// Communication API/Ethernet/API/bds_ethIPv4_setLocalIpAdr
///This function sets the IPv4 Address and Subnet Mask of the ECU.
///
///=======
/// Remarks:
///=======
///This function must be called from initialization task. 
///IP address shall be Unicast only. Multicast (from 0xE0000000 to 0xEFFFFFFF) or broadcast (0xFFFFFFFF) or 0 are not allowed.
///The Subnet mask(CIDR) can have any value from 1 to 31.
///If this API is called properly from OsIniProc(), then it will overwrite the IP address configured in easyConfig.
///The header file bds_ethIPv4_SetIPAdr.h shall be included for enabling usage of defines.
///----------
/// FFI:
///----------
///This API can be used in trusted partitions only. See Freedom from Interference (FFI) concept for more details.
///
///==================================================================		  	===================================================================================================
///Return value    								  							    Description
///==================================================================		  	===================================================================================================
///bds_ethIPv4_Adr_Mask_ok_E                                                    API call is successful
///bds_ethIPv4_Adr_Nok_E                                                        API call is invalid because of invalid IPv4 address, Unicast address expected.
///bds_ethIPv4_Mask_Nok_E 	                                                    API call is invalid because of invalid subnet mask, subnet mask should be 16.
///bds_ethIPv4_Api_NotAvailable_E                                               Not Available (e.g. busy, called too early in init, not called from OsIniProc etc.)
///
///==================================================================		   	===================================================================================================
///=======
///Code Example:
///=======
/// PROGRAM ETHERNET
/// VAR
///   bds_ethIPv4_Set_Adr_Mask_s1 : bds_ethIPv4_LocalIpAdr_ts;
///   flag_u8 : USINT := 0;
/// END_VAR
///
/// (* Set IP Address: 192.168.0.3 (0xC0A80003) *)
/// bds_ethIPv4_Set_Adr_Mask_s1.Ipv4Adr_u32 := 16#C0A80003; 
///
/// (* Set Subnet Mask: /16 (255.255.0.0) *)
/// bds_ethIPv4_Set_Adr_Mask_s1.Ipv4SubnetMask_u8 := 16;
///
/// (* Apply IP configuration *)
/// 
/// IF(flag_u8 = 0) THEN
/// bds_ethIPv4_setLocalIpAdr(bds_ethIPv4_Set_Adr_Mask_s1);
///
/// flag_u8 :=1;
/// END_IF
/// END_PROGRAM
///============================================================================
{attribute 'external_name' := 'cmp_rts_bds_ethIPv4_setLocalIpAdr'}
FUNCTION bds_ethIPv4_setLocalIpAdr : bds_ethIPv4_setLocalIpAdr_ts
VAR_INPUT
	//Data Structure for IPv4 Address and Subnet Mask
	bds_ethIPv4_setLocalIpAdr_s : bds_ethIPv4_LocalIpAdr_ts;
END_VAR

END_FUNCTION

// Communication API/Ethernet/API/bds_ethIPv4_getLocalIpAdr
///This function reads the IPv4 Address and Subnet Mask of the ECU.
///
///=======
/// Remarks:
///=======
///The header file bds_ethIPv4_SetIPAdr.h shall be included for enabling usage of defines.
///----------
/// FFI:
///----------
///This API can be used in trusted partitions only. See Freedom from Interference (FFI) concept for more details.
///
///==================================================================		  	===================================================================================================
///Return value    								  							    Description
///==================================================================		  	===================================================================================================
///bds_ethIPv4_Adr_Mask_ok_E                                                    API call is successful
///bds_ethIPv4_Api_NotAvailable_E                                               Not Available (e.g. busy, called too early in init, not called from OsIniProc etc.)
///bds_ethIPv4_NullPtr_E                                                        Invalid parameter passed
///==================================================================		   	===================================================================================================
///=======
///Code Example:
///=======
///PROGRAM ETHERNET
/// VAR
///    bds_ethIPv4_Get_Adr_Mask_s2 : bds_ethIPv4_LocalIpAdr_ts;
/// END_VAR
/// 
/// bds_ethIPv4_Get_Adr_Mask_s2.Ipv4Adr_u32 := 0;
/// bds_ethIPv4_Get_Adr_Mask_s2.Ipv4SubnetMask_u8 := 0;
///
/// bds_ethIPv4_getLocalIpAdr(ADR(bds_ethIPv4_Get_Adr_Mask_s2));
///
///END_PROGRAM
///============================================================================
{attribute 'external_name' := 'cmp_rts_bds_ethIPv4_getLocalIpAdr'}
FUNCTION bds_ethIPv4_getLocalIpAdr : bds_ethIPv4_getLocalIpAdr_ts
VAR_INPUT
	//Data Structure for IPv4 Address and Subnet Mask
	bds_ethIPv4_getLocalIpAdr_s : POINTER TO bds_ethIPv4_LocalIpAdr_ts;
END_VAR

END_FUNCTION

// Communication API/Ethernet/API/bds_ethIPv4_setDoipAdr
///This function configures the RC4x's and Tester's logical addresses for Diagnostic over IP (DoIP) communication. 
///
///=======
/// Remarks:
///=======
///This function shall be called from initialization task.
///The logical address of the RC4x (ecuLogAdr_u16) must fall within one of two valid ranges, as defined by ISO 13400-2:
/// Standard ECU addresses - 0x0001 to 0x0DFF
/// Extended ECU addresses - 0x1000 to 0x7FFF.
/// An address outside these ranges will result in bds_ethIPv4_retLogAdrNok_E.
///The Tester logical address (testerLogAdr_u16) must be within the range 0x0E00 to 0x0FFF. An address outside this range will result in bds_ethIPv4_retTesterAdrNok_E.
///If this API is not called, or called incorrectly (validation fails , bds_ethIPv4_retTesterAdrNok_E), the RC4x shall use the addresses from easyConfig.
///This function call overrides the statically configured values provided by easyConfig.
///----------
/// FFI:
///----------
///This API can be used in trusted partitions only. See Freedom from Interference (FFI) concept for more details.
///
///==================================================================		  	===================================================================================================
///Return value    								  							    Description
///==================================================================		  	===================================================================================================
///ecuLogAdr_u16                                                                API call is successful
///testerLogAdr_u16                                                             Tester logical address (valid range: 0x0E00-0x0FFF)
///
///==================================================================		   	===================================================================================================
///=======
///Code Example:
///=======
///PROGRAM ETHERNET
/// VAR
///    doipStatus : bds_ethIPv4_retDoipAdr_te;
///    flag_u8 : USINT := 0;
/// END_VAR

(* Configure ECU Logical Target Address and Tester Address Range
 *
 * ECU Logical Target Address = 0x0200
 * Tester Address Range Min   = 0x0E00
 *
 * NOTE: The Tester Address Range Max is internally defined in the stack.
 *)
/// IF(flag_u8 = 0) THEN
/// doipStatus := bds_ethIPv4_setDoipAdr(16#0200, 16#0E00);
/// 
/// flag_u8 := 1;
/// 
/// END_IF
///
(* Check return status *)
/// IF doipStatus = bds_ethIPv4_retAdrOk_E THEN
   (* DoIP address successfully configured*)
    
/// ELSE
    (* Error handling: DoIP address configuration failed*)
    
/// END_IF;

/// END_PROGRAM
///============================================================================
{attribute 'external_name' := 'cmp_rts_bds_ethIPv4_setDoipAdr'}
FUNCTION bds_ethIPv4_setDoipAdr : bds_ethIPv4_retDoipAdr_te
VAR_INPUT
	//RC4x logical address (valid ranges: 0x0001-0x0DFF or 0x1000-0x7FFF)
	ecuLogAdr_u16 : UINT;
	//Tester logical address (valid range: 0x0E00-0x0FFF)
	testerLogAdr_u16 : UINT;
END_VAR

END_FUNCTION

// Communication API/Ethernet/API/bds_ethIPv4_getLinkState
///This function returns the current physical link status of the RC4x's ethernet interface.
///
///=======
/// Remarks:
///=======
///This function provides the ethernet link status.
///----------
/// FFI:
///----------
///This API can be used in trusted partitions only. See Freedom from Interference (FFI) concept for more details.
///
///==================================================================		  	===================================================================================================
///Return value    								  							    Description
///==================================================================		  	===================================================================================================
///bds_ethIPv4_retLinkOk_E                                                      Link status retrieved successfully 
///bds_ethIPv4_retLinkNok_E                                                     Failed to get link status 
///bds_ethIPv4_retLinkNull_E                                                    Invalid parameter - NULL pointer passed as argument
///==================================================================		   	===================================================================================================
///=======
///Code Example:
///=======
/// PROGRAM ETHERNET
/// VAR
///    linkStateInfo_s : bds_ethIPv4_linkStateInfo_ts;
///    linkStatus_e : bds_ethIPv4_retlinkState_te;
/// END_VAR

/// Retrieve Ethernet link state
/// linkStatus_e := bds_ethIPv4_getLinkState(ADR(linkStateInfo_s));

/// IF linkStatus_e = bds_ethIPv4_retLinkOk_E THEN
    
///    IF linkStateInfo_s.currentState_e = bds_ethIPv4_linkUp_E THEN
///         Ethernet link is UP (normal communication possible)
        
///    ELSIF linkStateInfo_s.currentState_e = bds_ethIPv4_linkDown_E THEN
        (* Ethernet link is DOWN (no communication)
         Take fallback ACTION IF required*)
        
///    ELSE
        (* Link state is undefined (transitional or error state)*)
        
///    END_IF;
    
/// ELSE
    (* Error: Failed TO get link state
     Handle error CASE (e.g., LOG OR retry)*)
    
/// END_IF;

/// END_PROGRAM
///
///============================================================================
{attribute 'external_name' := 'cmp_rts_bds_ethIPv4_getLinkState'}
FUNCTION bds_ethIPv4_getLinkState : bds_ethIPv4_retLinkState_te
VAR_INPUT
  //A pointer to a bds_ethIPv4_linkStateInfo_ts structure. 
  //Upon execution, the currentState_e member of this structure will be updated with the current.
  //Ethernet link state (bds_ethIPv4_linkDown_E, bds_ethIPv4_linkUp_E, or bds_ethIPv4_linkUndef_E). 
  linkStateInfo_ps : POINTER TO bds_ethIPv4_linkStateInfo_ts;
END_VAR

END_FUNCTION

// Diagnostics API/UDS/API/bds_uds_setNodeIdTesterId
///This function sets the Node ID and Tester ID through Application Software (ASW) for the Bodas-Service instance.
///
///=======
/// Remarks:
///=======
///This function must be called from initialization task.  
///The header file bds_bsw.h shall be included for enabling usage of defines.
///To read the configured node ID and tester ID bds_uds_getNodeID can be used.
///BODAS-Service tool can't be used if Tester ID is set to other than 0xFA.
///
///
///===========
///ATTENTION
///===========
///The functional address is currently fixed to 0x18DBFFFA in the BODAS-Service tool. Communication will not work if the user modifies tester ID to other than 0xFA.
///It is recommended to use bds_uds_setNodeIdTesterId instead of bds_uds_updNodeIDinNVM.
///
///----------
/// FFI:
///----------
///This API can be used in trusted partitions only. See Freedom from Interference (FFI) concept for more details.
///
///==================================================================		  			===================================================================================================
///Return value    								  									    Description
///==================================================================		  			===================================================================================================
///bds_uds_nodeIdTesterIdOk_E															Node Id and Tester Id is set.
///bds_uds_nodeIdNotOk_E  																0xFF is broadcast node ID which cannot be used
///bds_uds_testerIdNotOk_E                                                              0xFF is broadcast tester ID which cannot be used 
///bds_uds_sameNodeIdTesterIdNotOk_E                                                    Node ID and tester ID value cannot be same. 
///bds_uds_setIDApiNotAvailable_E                                                       The API must be called from initialization task and cannot be called from elsewhere.
///
///==================================================================		   			===================================================================================================
///
///=======
///Code Example:
///=======
/// PROGRAM ETHERNET
/// VAR
///    return_e : bds_uds_setNodeIdTesterId_te;
///    flag_u8 : USINT :=0;
/// END_VAR
///
/// IF(flag_u8 = 0) THEN
/// return_e := bds_uds_setNodeIdTesterId(16#06, 16#08);
/// 
/// flag_u8 :=1;
/// END_IF
///
/// END_PROGRAM
///============================================================================
///
{attribute 'external_name' := 'cmp_rts_bds_uds_setNodeIdTesterId'}
FUNCTION bds_uds_setNodeIdTesterId : bds_uds_setNodeIdTesterId_te
VAR_INPUT
	//Node ID to be configured
	nodeId_u8 : USINT;
	//Tester ID to be configured
	testerId_u8 : USINT;
END_VAR

END_FUNCTION

// System API/SYS/API/bds_sys_regOverwriteOpHrsCbk
///This function bds_sys_regOverwriteOpHrsCbk() registers a callback function to replace the Environment data operating hours with customer-specific data.
///
///=======
/// Remarks:
///=======
///This function must be called from initialization task.
///If the bds_sys_regOverwriteOpHrs_pf callback is registered, Environment data operating hours will be updated from the callback implemented in ASW.
///If the bds_sys_regOverwriteOpHrs_pf callback is not registered, Environment data operating hours will be updated by BSW.
///This API allows customers to overwrite the ECU's operating hours with their preferred data, in the response to UDS service $1904.
///The size of customer specific data is 4 bytes.
///Operating hours cannot be changed. Only the time stamp that is stored with environmental data can be overwritten.
///
///----------
/// FFI:
///----------
///This API can be used in trusted partitions only. See Freedom from Interference (FFI) concept for more details.
///
///==================================================================		  		===================================================================================================
///Return value    								  									Description
///==================================================================		  		===================================================================================================
///bds_sys_regOpHrsOk_E																Callback function registered successfully 
///bds_sys_regOpHrsNullPtr_E                                                        A null pointer error occurred for the callback.
///bds_sys_regOpHrsApiNotAvailable_E                                                The API is only available from OsIniProc and cannot be called from elsewhere.
 
///==================================================================		   		===================================================================================================
///=======
///Code Example:
///=======
///
/// PROGRAM RegoverwriteOpHrs
/// VAR
///    bds_sys_regOverwriteOpHrs_ret : bds_sys_regOverwriteOpHrs_te; // Or appropriate enum type
///    flag_u8 : USINT := 0;
///
/// END_VAR
/// 
/// IF (flag_u8 = 0)THEN
///
/// bds_sys_regOverwriteOpHrs_ret := bds_sys_regOverwriteOpHrsCbk(bds_sys_OverWrtED_pf);
/// flag_u8 :=1;
/// 
/// END_IF
///
/// FUNCTION bds_sys_OverWrtED_pf
/// VAR_INPUT
///    ED_Value_32_ptr : POINTER TO UDINT; // Pointer to uint32
/// END_VAR
///
/// ED_Value_32_ptr^ := 16#400;
///
///============================================================================
{attribute 'external_name' := 'cmp_rts_bds_sys_regOverwriteOpHrsCbk'}
FUNCTION bds_sys_regOverwriteOpHrsCbk : bds_sys_regOverwriteOpHrs_te
VAR_INPUT
	bds_sys_regOverwriteOpHrs_pf : UINT;
END_VAR

END_FUNCTION

// System API/SYS/API/bds_codesys_setForcingWritingMode
{attribute 'external_name' := 'cmp_rts_bds_codesys_setForcingWritingMode'}
///This function is used to enable/disable forcing and writing feature inside CODESYS IDE
///
///----------
/// FFI:
///----------
///This API can be used in trusted partitions only. See Freedom from Interference (FFI) concept for more details.
///
///----------
/// DANGER:
///----------
///
///Software running on the ECU can be manipulated with forcing or writing. That will lead to both a security and a safety risk. Life and health can be endangered. Thus, it must be impossible to use forcing or writing on serial machines.
///
///
///==================================================================		  			===================================================================================================
///Return value    								  									Description
///==================================================================		  			===================================================================================================
///None																				None
///
///==================================================================		   			===================================================================================================
///
///
///=======
///Code Example:
///=======
///============================================================================
///
///PROGRAM PLC_PRG
///  VAR
///  
///  END_VAR
///
///  (* Enable Forcing and Writing *)
///  
///  bds_codesys_setForcingWritingMode(16#FFFF);
///
///============================================================================
FUNCTION bds_codesys_setForcingWritingMode
VAR_INPUT
		///Indicates whether Forcing and Writing should be enabled or disabled.
	///
	///Possible values:
	///    + BDS_DISABLE_FORCINGWRITING_DU16 (16#0000)           : Disable Forcing and Writing.
	///    + BDS_ENABLE_FORCINGWRITING_DU16  (16#FFFF)           : Enable Forcing and Writing.
	mode_u16: UINT;
END_VAR

END_FUNCTION
